// TIA Portal V19 export
VAR_GLOBAL   // PLC tag table "Servo"
   DI_ServoHomming AT %I8.2 : Bool;
END_VAR
